(* IEC 61131-3 sources: SortJet_MasterSPS_Aufbau.fbsproj/11_MMI_Kommunikation/IoControl, 10 files *)

(* ---- GetBitStatus.fn.st ---- *)
(* METADATA
{
	"v3Meta": {
		"objectGuid": "3b6ea6e4-8fcd-474b-9f1e-9c8a8e0a159e"
	}
}
*)
FUNCTION GetBitStatus : BOOL
VAR_INPUT
  wpWatchIoNr : WORD;
END_VAR
VAR
  wlByteIndex : WORD;
  wlBitIndex : WORD;
  uclRet   : BYTE;
  ucpValue : BYTE;
END_VAR
wlByteIndex := wpWatchIoNr / 8;
wlBitIndex  := wpWatchIoNr MOD 8;

ucpValue := TCPMain.l_fb_SortjetHMI.SpsToMmi.aucControlSystem[ wlByteIndex ];

uclRet := ucpValue;

CASE wlBitIndex OF

  0: GetBitStatus := uclRet.0;

  1: GetBitStatus := uclRet.1;

  2: GetBitStatus := uclRet.2;

  3: GetBitStatus := uclRet.3;

  4: GetBitStatus := uclRet.4;

  5: GetBitStatus := uclRet.5;

  6: GetBitStatus := uclRet.6;

  7: GetBitStatus := uclRet.7;

END_CASE
END_FUNCTION

(* ---- ResetIoControl.fn.st ---- *)
(* METADATA
{
	"v3Meta": {
		"objectGuid": "57b43017-bb28-437d-982e-b60f799a1ca9"
	}
}
*)
FUNCTION ResetIoControl : BOOL
VAR_INPUT
  wpControlIndex : WORD;
END_VAR
VAR
  wlByteIndex : WORD;
  wlBitIndex  : WORD;
  ucValue     : BYTE;
END_VAR

wlByteIndex := wpControlIndex / 8;
wlBitIndex  := wpControlIndex MOD 8;

// Überwachung deaktivieren
aicgIoControl[ wpControlIndex ].tWatchStart := T#0ms;

// Meldungsbit zurücksetzen
ucValue := TCPMain.l_fb_SortjetHMI.SpsToMmi.aucControlSystem[ wlByteIndex ];
ucValue := SetBitStatus( ucValue, wlBitIndex, FALSE );
TCPMain.l_fb_SortjetHMI.SpsToMmi.aucControlSystem[ wlByteIndex ] := ucValue;
END_FUNCTION

(* ---- SetBitStatus.fn.st ---- *)
(* METADATA
{
	"v3Meta": {
		"objectGuid": "e3d893c7-2aa8-4b16-bd4f-cc2db28304fb"
	}
}
*)
FUNCTION SetBitStatus : BYTE
VAR_INPUT
  ucpValue : BYTE;
  wpBitPos : WORD;
  bpStatus : BOOL;
END_VAR
VAR
  uclRet : BYTE;
END_VAR
// Bit in eine Word setzen
uclRet := ucpValue;

CASE wpBitPos OF

  0:uclRet.0  := bpStatus;

  1:uclRet.1  := bpStatus;

  2:uclRet.2  := bpStatus;

  3:uclRet.3  := bpStatus;

  4:uclRet.4  := bpStatus;

  5:uclRet.5  := bpStatus;

  6:uclRet.6  := bpStatus;

  7:uclRet.7  := bpStatus;

END_CASE

SetBitStatus := uclRet;
END_FUNCTION

(* ---- SetIoControl.fn.st ---- *)
(* METADATA
{
	"v3Meta": {
		"objectGuid": "cdf47146-760f-48c9-a8df-c674983d5b70"
	}
}
*)
FUNCTION SetIoControl : BOOL
VAR_INPUT
  wpControlIndex : WORD;
END_VAR
VAR
  wlByteIndex : WORD;
  wlBitIndex  : WORD;
  ucValue     : BYTE;
END_VAR

wlByteIndex := wpControlIndex / 8;
wlBitIndex  := wpControlIndex MOD 8;

ucValue := TCPMain.l_fb_SortjetHMI.SpsToMmi.aucControlSystem[ wlByteIndex ];

ucValue := SetBitStatus( ucValue, wlBitIndex, TRUE );

TCPMain.l_fb_SortjetHMI.SpsToMmi.aucControlSystem[ wlByteIndex ] := ucValue;

SetIoControl := TRUE;
END_FUNCTION

(* ---- SpsError.fn.st ---- *)
(* METADATA
{
	"v3Meta": {
		"objectGuid": "8b5c3fca-ed53-4ab3-83d7-c24b940f4322"
	}
}
*)
FUNCTION SpsError : BOOL
VAR_INPUT
  wpFehlerGruppe    : WORD;
  wpErrorNr         : WORD;
  wpStationsnummmer : WORD;
  wpAutomatikkreis  : WORD;
  awpDaten          : ARRAY [0..25] OF WORD;
END_VAR
VAR
  smlMessage : SpsMessage;
END_VAR

smlMessage.wAuftrag := SB0_SPS_ERROR;

smlMessage.awDaten[0] := HMI_GetWORD(ADR(wpFehlerGruppe));
smlMessage.awDaten[1] := HMI_GetWORD(ADR(wpErrorNr));
smlMessage.awDaten[2] := HMI_GetWORD(ADR(wpStationsnummmer));
smlMessage.awDaten[3] := HMI_GetWORD(ADR(wpAutomatikkreis));

HMI_PutWORD( pbyAddr := ADR( smlMessage.awDaten ) + 8  , wVal := awpDaten[0] );
HMI_PutWORD( pbyAddr := ADR( smlMessage.awDaten ) + 10 , wVal := awpDaten[1] );
HMI_PutWORD( pbyAddr := ADR( smlMessage.awDaten ) + 12 , wVal := awpDaten[2] );
HMI_PutWORD( pbyAddr := ADR( smlMessage.awDaten ) + 14 , wVal := awpDaten[3] );
HMI_PutWORD( pbyAddr := ADR( smlMessage.awDaten ) + 16 , wVal := awpDaten[4] );
HMI_PutWORD( pbyAddr := ADR( smlMessage.awDaten ) + 18 , wVal := awpDaten[5] );
HMI_PutWORD( pbyAddr := ADR( smlMessage.awDaten ) + 20 , wVal := awpDaten[6] );
HMI_PutWORD( pbyAddr := ADR( smlMessage.awDaten ) + 22 , wVal := awpDaten[7] );
HMI_PutWORD( pbyAddr := ADR( smlMessage.awDaten ) + 24 , wVal := awpDaten[8] );
HMI_PutWORD( pbyAddr := ADR( smlMessage.awDaten ) + 26 , wVal := awpDaten[9] );
HMI_PutWORD( pbyAddr := ADR( smlMessage.awDaten ) + 28 , wVal := awpDaten[10] );
HMI_PutWORD( pbyAddr := ADR( smlMessage.awDaten ) + 30 , wVal := awpDaten[11] );
HMI_PutWORD( pbyAddr := ADR( smlMessage.awDaten ) + 32 , wVal := awpDaten[12] );
HMI_PutWORD( pbyAddr := ADR( smlMessage.awDaten ) + 34 , wVal := awpDaten[13] );
HMI_PutWORD( pbyAddr := ADR( smlMessage.awDaten ) + 36 , wVal := awpDaten[14] );
HMI_PutWORD( pbyAddr := ADR( smlMessage.awDaten ) + 38 , wVal := awpDaten[15] );
HMI_PutWORD( pbyAddr := ADR( smlMessage.awDaten ) + 40 , wVal := awpDaten[16] );
HMI_PutWORD( pbyAddr := ADR( smlMessage.awDaten ) + 42 , wVal := awpDaten[17] );
HMI_PutWORD( pbyAddr := ADR( smlMessage.awDaten ) + 44 , wVal := awpDaten[18] );
HMI_PutWORD( pbyAddr := ADR( smlMessage.awDaten ) + 46 , wVal := awpDaten[19] );
HMI_PutWORD( pbyAddr := ADR( smlMessage.awDaten ) + 48 , wVal := awpDaten[20] );
HMI_PutWORD( pbyAddr := ADR( smlMessage.awDaten ) + 50 , wVal := awpDaten[21] );
HMI_PutWORD( pbyAddr := ADR( smlMessage.awDaten ) + 52 , wVal := awpDaten[22] );
HMI_PutWORD( pbyAddr := ADR( smlMessage.awDaten ) + 54 , wVal := awpDaten[23] );
HMI_PutWORD( pbyAddr := ADR( smlMessage.awDaten ) + 56 , wVal := awpDaten[24] );
HMI_PutWORD( pbyAddr := ADR( smlMessage.awDaten ) + 58 , wVal := awpDaten[25] );

TCPMain.l_fb_SortjetHMI.PutMsg( smpSpsMessage := smlMessage, bpTrig := FALSE );
END_FUNCTION

(* ---- SpsHinweis.fn.st ---- *)
(* METADATA
{
	"v3Meta": {
		"objectGuid": "5fb299a3-7eb3-4628-8413-c7458efde9d6"
	}
}
*)
FUNCTION SpsHinweis : BOOL
VAR_INPUT
  wpFehlerGruppe    : WORD;
  wpErrorNr         : WORD;
  wpStationsnummmer : WORD;
  wpAutomatikkreis  : WORD;
  awpDaten          : ARRAY [0..25] OF WORD;
END_VAR
VAR
  smlMessage : SpsMessage;
END_VAR

smlMessage.wAuftrag := SB0_SPS_HINWEIS;

smlMessage.awDaten[0] := HMI_GetWORD(ADR(wpFehlerGruppe));
smlMessage.awDaten[1] := HMI_GetWORD(ADR(wpErrorNr));
smlMessage.awDaten[2] := HMI_GetWORD(ADR(wpStationsnummmer));
smlMessage.awDaten[3] := HMI_GetWORD(ADR(wpAutomatikkreis));

HMI_PutWORD( pbyAddr := ADR( smlMessage.awDaten ) + 8  , wVal := awpDaten[0] );
HMI_PutWORD( pbyAddr := ADR( smlMessage.awDaten ) + 10 , wVal := awpDaten[1] );
HMI_PutWORD( pbyAddr := ADR( smlMessage.awDaten ) + 12 , wVal := awpDaten[2] );
HMI_PutWORD( pbyAddr := ADR( smlMessage.awDaten ) + 14 , wVal := awpDaten[3] );
HMI_PutWORD( pbyAddr := ADR( smlMessage.awDaten ) + 16 , wVal := awpDaten[4] );
HMI_PutWORD( pbyAddr := ADR( smlMessage.awDaten ) + 18 , wVal := awpDaten[5] );
HMI_PutWORD( pbyAddr := ADR( smlMessage.awDaten ) + 20 , wVal := awpDaten[6] );
HMI_PutWORD( pbyAddr := ADR( smlMessage.awDaten ) + 22 , wVal := awpDaten[7] );
HMI_PutWORD( pbyAddr := ADR( smlMessage.awDaten ) + 24 , wVal := awpDaten[8] );
HMI_PutWORD( pbyAddr := ADR( smlMessage.awDaten ) + 26 , wVal := awpDaten[9] );
HMI_PutWORD( pbyAddr := ADR( smlMessage.awDaten ) + 28 , wVal := awpDaten[10] );
HMI_PutWORD( pbyAddr := ADR( smlMessage.awDaten ) + 30 , wVal := awpDaten[11] );
HMI_PutWORD( pbyAddr := ADR( smlMessage.awDaten ) + 32 , wVal := awpDaten[12] );
HMI_PutWORD( pbyAddr := ADR( smlMessage.awDaten ) + 34 , wVal := awpDaten[13] );
HMI_PutWORD( pbyAddr := ADR( smlMessage.awDaten ) + 36 , wVal := awpDaten[14] );
HMI_PutWORD( pbyAddr := ADR( smlMessage.awDaten ) + 38 , wVal := awpDaten[15] );
HMI_PutWORD( pbyAddr := ADR( smlMessage.awDaten ) + 40 , wVal := awpDaten[16] );
HMI_PutWORD( pbyAddr := ADR( smlMessage.awDaten ) + 42 , wVal := awpDaten[17] );
HMI_PutWORD( pbyAddr := ADR( smlMessage.awDaten ) + 44 , wVal := awpDaten[18] );
HMI_PutWORD( pbyAddr := ADR( smlMessage.awDaten ) + 46 , wVal := awpDaten[19] );
HMI_PutWORD( pbyAddr := ADR( smlMessage.awDaten ) + 48 , wVal := awpDaten[20] );
HMI_PutWORD( pbyAddr := ADR( smlMessage.awDaten ) + 50 , wVal := awpDaten[21] );
HMI_PutWORD( pbyAddr := ADR( smlMessage.awDaten ) + 52 , wVal := awpDaten[22] );
HMI_PutWORD( pbyAddr := ADR( smlMessage.awDaten ) + 54 , wVal := awpDaten[23] );
HMI_PutWORD( pbyAddr := ADR( smlMessage.awDaten ) + 56 , wVal := awpDaten[24] );
HMI_PutWORD( pbyAddr := ADR( smlMessage.awDaten ) + 58 , wVal := awpDaten[25] );

TCPMain.l_fb_SortjetHMI.PutMsg( smpSpsMessage := smlMessage, bpTrig := FALSE );
END_FUNCTION

(* ---- SpsLogString.fn.st ---- *)
(* METADATA
{
	"v3Meta": {
		"objectGuid": "3382b282-4d75-484e-8f31-3dfec2faf444"
	}
}
*)
FUNCTION SpsLogString : BOOL
VAR_INPUT
  spLogString : STRING(59);
END_VAR
VAR
  smlMessage     : SpsMessage;
  i,j            : WORD;
END_VAR

smlMessage.wAuftrag := SB0_SPS_LOGSTRING;

i:=SIZEOF(spLogString);
j:=SIZEOF(smlMessage.awDaten);

SysMemCpy( ADR( smlMessage.awDaten ), ADR( spLogString ), SIZEOF(spLogString) );

TCPMain.l_fb_SortjetHMI.PutMsg( smpSpsMessage := smlMessage, bpTrig := FALSE );
END_FUNCTION

(* ---- SpsWarnung.fn.st ---- *)
(* METADATA
{
	"v3Meta": {
		"objectGuid": "7de6b20f-9c42-4ee5-9d4c-1f3931e72fe6"
	}
}
*)
FUNCTION SpsWarnung : BOOL
VAR_INPUT
  wpFehlerGruppe    : WORD;
  wpErrorNr         : WORD;
  wpStationsnummmer : WORD;
  wpAutomatikkreis  : WORD;
  awpDaten          : ARRAY [0..25] OF WORD;
END_VAR
VAR
  smlMessage : SpsMessage;
END_VAR

smlMessage.wAuftrag := SB0_SPS_WARNUNG;

smlMessage.awDaten[0] := HMI_GetWORD(ADR(wpFehlerGruppe));
smlMessage.awDaten[1] := HMI_GetWORD(ADR(wpErrorNr));
smlMessage.awDaten[2] := HMI_GetWORD(ADR(wpStationsnummmer));
smlMessage.awDaten[3] := HMI_GetWORD(ADR(wpAutomatikkreis));

HMI_PutWORD( pbyAddr := ADR( smlMessage.awDaten ) + 8  , wVal := awpDaten[0] );
HMI_PutWORD( pbyAddr := ADR( smlMessage.awDaten ) + 10 , wVal := awpDaten[1] );
HMI_PutWORD( pbyAddr := ADR( smlMessage.awDaten ) + 12 , wVal := awpDaten[2] );
HMI_PutWORD( pbyAddr := ADR( smlMessage.awDaten ) + 14 , wVal := awpDaten[3] );
HMI_PutWORD( pbyAddr := ADR( smlMessage.awDaten ) + 16 , wVal := awpDaten[4] );
HMI_PutWORD( pbyAddr := ADR( smlMessage.awDaten ) + 18 , wVal := awpDaten[5] );
HMI_PutWORD( pbyAddr := ADR( smlMessage.awDaten ) + 20 , wVal := awpDaten[6] );
HMI_PutWORD( pbyAddr := ADR( smlMessage.awDaten ) + 22 , wVal := awpDaten[7] );
HMI_PutWORD( pbyAddr := ADR( smlMessage.awDaten ) + 24 , wVal := awpDaten[8] );
HMI_PutWORD( pbyAddr := ADR( smlMessage.awDaten ) + 26 , wVal := awpDaten[9] );
HMI_PutWORD( pbyAddr := ADR( smlMessage.awDaten ) + 28 , wVal := awpDaten[10] );
HMI_PutWORD( pbyAddr := ADR( smlMessage.awDaten ) + 30 , wVal := awpDaten[11] );
HMI_PutWORD( pbyAddr := ADR( smlMessage.awDaten ) + 32 , wVal := awpDaten[12] );
HMI_PutWORD( pbyAddr := ADR( smlMessage.awDaten ) + 34 , wVal := awpDaten[13] );
HMI_PutWORD( pbyAddr := ADR( smlMessage.awDaten ) + 36 , wVal := awpDaten[14] );
HMI_PutWORD( pbyAddr := ADR( smlMessage.awDaten ) + 38 , wVal := awpDaten[15] );
HMI_PutWORD( pbyAddr := ADR( smlMessage.awDaten ) + 40 , wVal := awpDaten[16] );
HMI_PutWORD( pbyAddr := ADR( smlMessage.awDaten ) + 42 , wVal := awpDaten[17] );
HMI_PutWORD( pbyAddr := ADR( smlMessage.awDaten ) + 44 , wVal := awpDaten[18] );
HMI_PutWORD( pbyAddr := ADR( smlMessage.awDaten ) + 46 , wVal := awpDaten[19] );
HMI_PutWORD( pbyAddr := ADR( smlMessage.awDaten ) + 48 , wVal := awpDaten[20] );
HMI_PutWORD( pbyAddr := ADR( smlMessage.awDaten ) + 50 , wVal := awpDaten[21] );
HMI_PutWORD( pbyAddr := ADR( smlMessage.awDaten ) + 52 , wVal := awpDaten[22] );
HMI_PutWORD( pbyAddr := ADR( smlMessage.awDaten ) + 54 , wVal := awpDaten[23] );
HMI_PutWORD( pbyAddr := ADR( smlMessage.awDaten ) + 56 , wVal := awpDaten[24] );
HMI_PutWORD( pbyAddr := ADR( smlMessage.awDaten ) + 58 , wVal := awpDaten[25] );

TCPMain.l_fb_SortjetHMI.PutMsg( smpSpsMessage := smlMessage, bpTrig := FALSE );
END_FUNCTION

(* ---- WatchIo.fn.st ---- *)
(* METADATA
{
	"v3Meta": {
		"objectGuid": "9bbc4f4b-7c56-4bbd-9f87-a841e4609bac"
	}
}
*)
FUNCTION WatchIo : BOOL
VAR_INPUT
  bpStatus : BOOL;
  wpControlIndex : WORD;
END_VAR
VAR
  wlByteIndex : WORD;
  wlBitIndex  : WORD;
  ucValue     : BYTE;
END_VAR
IF NOT bgDeaktiviereWatchIOs THEN
  IF bpStatus <> GetBitStatus(wpControlIndex) THEN
    wlByteIndex := wpControlIndex / 8;
    wlBitIndex  := wpControlIndex MOD 8;
    // Meldungsbit zurücksetzen
    ucValue := TCPMain.l_fb_SortjetHMI.SpsToMmi.aucControlSystem[ wlByteIndex ];
    IF bpStatus THEN
      ucValue := SetBitStatus( ucValue, wlBitIndex, TRUE );
    ELSE
      aicgIoControl[ wpControlIndex ].tWatchStart := T#0MS;
      ucValue := SetBitStatus( ucValue, wlBitIndex, FALSE );
    END_IF
    TCPMain.l_fb_SortjetHMI.SpsToMmi.aucControlSystem[ wlByteIndex ] := ucValue;
  END_IF
END_IF
END_FUNCTION

(* ---- WatchIoControl.fn.st ---- *)
(* METADATA
{
	"v3Meta": {
		"objectGuid": "8ac789ad-b8f8-4460-adb8-3fa1c010b792"
	}
}
*)
FUNCTION WatchIoControl : BOOL
VAR_INPUT
  tpTimeOut      : TIME;
  wpControlIndex : WORD;
  bpStatus       : BOOL;
END_VAR
VAR
  blResult    : BOOL;
  tlLaufzeit  : TIME;
END_VAR

blResult := FALSE;

IF NOT bgDeaktiviereWatchIOs THEN
  aicgIoControl[ wpControlIndex ].tTimeOut := tpTimeOut;
  IF bpStatus THEN
    IF( aicgIoControl[ wpControlIndex ].tWatchStart > T#0ms )THEN

      tlLaufzeit := TIME() - aicgIoControl[ wpControlIndex ].tWatchStart;

      IF( tlLaufzeit >= aicgIoControl[ wpControlIndex ].tTimeOut )THEN
        SetIoControl( wpControlIndex );
        blResult := TRUE;
      END_IF

    ELSE
      // Überwachung starten
      aicgIoControl[ wpControlIndex ].tWatchStart := TIME();
    END_IF
  ELSE
    ResetIoControl( wpControlIndex := wpControlIndex );
  END_IF

END_IF

WatchIoControl := blResult;
END_FUNCTION
